Fanuc KAREL source: kc00022.KL

-- PROVISIONAL review KL for V940-1; original PC SHA256 718d1be86ac7a8c76f165ae822f29442c6c4509c1d331afd5b0aa397a3469608
-- Incomplete behavior may be omitted. Consult companion uncertainty JSON. Do not deploy.
PROGRAM KC00022
%NOLOCKGROUP
BEGIN
  -- V9_ZERO_TABLE_METADATA_HINT layout=0002_ascii; no indexed target words; source/name/runtime held
  -- UNRESOLVED_PC offsets 5-22; opcodes 3F,75
  -- UNRESOLVED_PC offsets 27-45; opcodes 27,22,2A,22,31
  -- UNRESOLVED_PC offsets 50-54; opcodes 7F
END KC00022
